// TIA Portal project "PLC_hackathon_2026_V21" (V21)

(* hardware
DEVICE "S71500/ET200MP station_1"  S7-1500 station
   slot 0: "Rail_0"  Rack  6ES7 590-1***0-0AA0
   slot 1: "PLC_1"  CPU 1515-2 PN  6ES7 515-2AM01-0AB0  V2.6
      slot 3: "CPU display_1"  6ES7591-1BA00-0AA0
DEVICE "PC-System_1"  SIMATIC PC station
   slot 0: "SIMATIC PC station"  Rail  SIMATIC PC-Station  V1.0
      slot 125: "Stationmanager"  Station_Manager  V6.0.4
   slot 1: "HMI_RT_1"  WinCC RT Advanced  6AV2 104-0xxxx-xxxx  17.0.0.0
      slot 33792: "Host interface"  Host interface
   slot 2: "IE general_1"  IE General  IE_CP  V8.2.0
*)

// ===== PLC "PLC_1"  CPU 1515-2 PN =====
// protected blocks, not shown: "Crane_manipulation"

VAR_GLOBAL   // PLC tag table "Default tag table"
   "x_position" AT %MB104 : SInt;
   "y_position" AT %MB105 : SInt;
   "bay_ID" AT %MB106 : USInt;
   "number_of_manipulations" AT %MD107 : UDInt;
   "time" AT %MD112 : Real;
END_VAR

VAR_GLOBAL   // PLC tag table "Crane_command"
   "new_x_position" AT %MB100 : SInt;   // X position for the move command
   "new_y_position" AT %MB101 : SInt;   // Y position for the move command
   "new_bay_ID" AT %MB102 : USInt;   // Bay ID for the move command
   "new_command_ID" AT %MB103 : USInt;   // ID of the command
END_VAR

DATA_BLOCK "Current_state_of_Bay0"   // DB10
{ S7_Optimized_Access := 'TRUE' }
VERSION : 0.1
   VAR
      Bay0 : Array[0..3, 0..11] of UInt;
   END_VAR
BEGIN
   Bay0[0,0] := 123;
   Bay0[0,1] := 326;
   Bay0[0,2] := 987;
END_DATA_BLOCK

DATA_BLOCK "Current_state_of_Bay1"   // DB11
{ S7_Optimized_Access := 'TRUE' }
VERSION : 0.1
   VAR
      Bay1 : Array[0..3, 0..11] of UInt;
   END_VAR
BEGIN
   Bay1[0,1] := 246;
   Bay1[0,7] := 675;
   Bay1[1,5] := 777;
END_DATA_BLOCK

DATA_BLOCK "From_Bay0_to_Bay1"   // DB20
{ S7_Optimized_Access := 'TRUE' }
VERSION : 0.1
   VAR
      IDs_of_the_containers : Array[1..48] of UInt;
   END_VAR
BEGIN
   IDs_of_the_containers[12] := 0;
   IDs_of_the_containers[18] := 0;
   IDs_of_the_containers[4] := 444;
   IDs_of_the_containers[1] := 111;
   IDs_of_the_containers[2] := 222;
   IDs_of_the_containers[3] := 333;
   IDs_of_the_containers[5] := 555;
   IDs_of_the_containers[6] := 666;
   IDs_of_the_containers[7] := 777;
END_DATA_BLOCK

DATA_BLOCK "From_Bay1_to_Bay0"   // DB21
{ S7_Optimized_Access := 'TRUE' }
VERSION : 0.1
   VAR
      Bay1_IDs_of_the_containers : Array[1..48] of UInt;
   END_VAR
BEGIN
   Bay1_IDs_of_the_containers[15] := 0;
   Bay1_IDs_of_the_containers[22] := 0;
   Bay1_IDs_of_the_containers[1] := 123;
   Bay1_IDs_of_the_containers[2] := 124;
   Bay1_IDs_of_the_containers[3] := 125;
END_DATA_BLOCK

// folder: Constants

DATA_BLOCK "Global_constants"   // DB1
{ S7_Optimized_Access := 'TRUE' }
VERSION : 0.1
   VAR
      container_width_in_m : Real := 2.3;   // Container width in meters
      container_length_in_m : Real := 6.0;   // Container length in meters
      velocity_of_the_crane_in_m_per_s : Real := 1.0;   // Velocity of the crane in meters per second
      time_to_lift_a_container_in_s : Real := 20.0;   // Time needed to lower the hook, hook up a container and lift it in seconds
      time_to_put_down_a_container_in_s : Real := 20.0;   // Time needed to put down a container, release it, and lift up the hook in seconds
   END_VAR
BEGIN
END_DATA_BLOCK

// folder: (top level)

ORGANIZATION_BLOCK "Cyclic interrupt"   // OB30, LAD, CyclicInterrupt
{ S7_Optimized_Access := 'TRUE' }
VERSION : 0.1
   VAR_INPUT
      Initial_Call : Bool;   // Initial call of this OB
      Event_Count : Int;   // Events discarded
   END_VAR
BEGIN

REGION Network 1: Crane manipulation
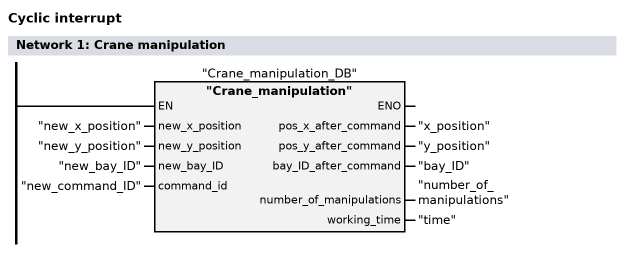
   RUNG wire#powerrail
      "Crane_manipulation_DB"(new_x_position := "new_x_position", new_y_position := "new_y_position", new_bay_ID := "new_bay_ID", command_id := "new_command_ID", pos_x_after_command => "x_position", pos_y_after_command => "y_position", bay_ID_after_command => "bay_ID", number_of_manipulations => "number_of_manipulations", working_time => "time")
   END_RUNG
   // the same network as SCL:
   "Crane_manipulation_DB"(new_x_position := "new_x_position",   // "Crane_manipulation"
                           new_y_position := "new_y_position",
                           new_bay_ID := "new_bay_ID",
                           command_id := "new_command_ID",
                           pos_x_after_command => "x_position",
                           pos_y_after_command => "y_position",
                           bay_ID_after_command => "bay_ID",
                           number_of_manipulations => "number_of_manipulations",
                           working_time => "time");
END_REGION
END_ORGANIZATION_BLOCK

ORGANIZATION_BLOCK "Startup"   // OB100, SCL, Startup
TITLE = "Complete Restart"
{ S7_Optimized_Access := 'TRUE' }
VERSION : 0.1
   VAR_INPUT
      LostRetentive : Bool;   // True if retentive data are lost
      LostRTC : Bool;   // True if date and time are lost
   END_VAR
BEGIN
   // define the inital state of the shipyard
   "Crane_manipulation_DB".command_id := 0; // set "do nothing" command
   "Crane_manipulation_DB".current_bay_ID := 1; // the crane starting bay ID set to 1 (left of the ship)
   "Crane_manipulation_DB".current_x_position_in_bay := 0; // starting X position of the crane
   "Crane_manipulation_DB".current_y_position_in_bay := 0; // starting Y position of the crane

   //define startup command parameters
   "new_x_position" := 0; // starting X position of the crane
   "new_y_position" := 0; // starting Y position of the crane
   "new_bay_ID" := 1; // the crane starting bay ID set to 1 (left of the ship)
   "new_command_ID" := 0; // set "do nothing" command

   // reset of evaluation parameters
   "Crane_manipulation_DB".total_number_of_manipulations := 0; // reset total number of the crane manipulations
   "Crane_manipulation_DB".total_time := 0.0; // reset of total time
END_ORGANIZATION_BLOCK

(* ===== HMI "HMI_RT_1" =====
connection "HMI_Connection_1": ETHERNET, S7_1500_OMS

HMI tags "Default tag table"
   "time" : Real = PLC time AT %MD112, 1 s

screen "Screen_1" 1024x768
   TextField "Text field_1" at 20,17 size 95x22; Text 'PLC+ 2019:'
   IOField "I/O field_1" at 86,66 size 96x32; FormatPattern s999999999.999
      ProcessValue <- "time"
*)